Fanuc KAREL source: kt00106.KL

-- PROVISIONAL review KL for V1013-1; original PC SHA256 6ff60232844880fed4de48d1acf513a84916199fc54f7c6ee0a3c9b76619d910
-- Incomplete behavior may be omitted. Consult companion uncertainty JSON. Do not deploy.
PROGRAM KT00106
%NOLOCKGROUP
VAR
  R1 : REAL
  I2 : INTEGER
  OUT : REAL
BEGIN
  -- UNRESOLVED_PC offsets 5-16; opcodes 2E,23
  -- UNRESOLVED_PC offsets 21-32; opcodes 2E,23
  -- UNRESOLVED_PC offsets 37-57; opcodes 21,21,64,6C,23
  -- UNRESOLVED_PC offsets 62-66; opcodes 7F
END KT00106
